// TIA Portal V19 export
VAR_GLOBAL   // PLC tag table "R3_IN"
   "ByteIN :0 R3" AT %IB154 : Byte;   // System Bits 1
   "ByteIN :1 R3" AT %IB155 : Byte;   // System Bits 2
   "ByteIN :2 R3" AT %IB156 : Byte;   // Signals
   "ByteIN :3 R3" AT %IB157 : Byte;   // Signals
   "ByteIN :4 R3" AT %IB158 : Byte;   // CMD
   "ByteIN :5 R3" AT %IB159 : Byte;
   "ByteIN :6 R3" AT %IB160 : Byte;
   "ByteIN :7 R3" AT %IB161 : Byte;
   "ByteIN :8 R3" AT %IB162 : Byte;
   "ByteIN :9 R3" AT %IB163 : Byte;
   "ByteIN :10 R3" AT %IB164 : Byte;
   "ByteIN :11 R3" AT %IB165 : Byte;
   "ByteIN :12 R3" AT %IB166 : Byte;
   "ByteIN :13 R3" AT %IB167 : Byte;
   "ByteIN :14 R3" AT %IB168 : Byte;
   "ByteIN :15 R3" AT %IB169 : Byte;
   "ByteIN :16 R3" AT %IB170 : Byte;
   "ByteIN :17 R3" AT %IB171 : Byte;
   "ByteIN :18 R3" AT %IB172 : Byte;
   "ByteIN :19 R3" AT %IB173 : Byte;
   "ByteIN :20 R3" AT %IB174 : Byte;
   "ByteIN :21 R3" AT %IB175 : Byte;
   "ByteIN :22 R3" AT %IB176 : Byte;
   "ByteIN :23 R3" AT %IB177 : Byte;
   "ByteIN :24 R3" AT %IB178 : Byte;
   "ByteIN :25 R3" AT %IB179 : Byte;
   "ByteIN :26 R3" AT %IB180 : Byte;
   "ByteIN :27 R3" AT %IB181 : Byte;
   "ByteIN :28 R3" AT %IB182 : Byte;
   "ByteIN :29 R3" AT %IB183 : Byte;
   "ByteIN :30 R3" AT %IB184 : Byte;
   "ByteIN :31 R3" AT %IB185 : Byte;
   "ByteIN :32 R3" AT %IB186 : Byte;
   "ByteIN :33 R3" AT %IB187 : Byte;
   "ByteIN :34 R3" AT %IB188 : Byte;
   "ByteIN :35 R3" AT %IB189 : Byte;
   "ByteIN :36 R3" AT %IB190 : Byte;
   "ByteIN :37 R3" AT %IB191 : Byte;
   "ByteIN :38 R3" AT %IB192 : Byte;
   "ByteIN :39 R3" AT %IB193 : Byte;
   "ByteIN :40 R3" AT %IB194 : Byte;
   "ByteIN :41 R3" AT %IB195 : Byte;
   "ByteIN :42 R3" AT %IB196 : Byte;
   "ByteIN :43 R3" AT %IB197 : Byte;
   "ByteIN :44 R3" AT %IB198 : Byte;
   "ByteIN :45 R3" AT %IB199 : Byte;
   "ByteIN :46 R3" AT %IB200 : Byte;
   "ByteIN :47 R3" AT %IB201 : Byte;
   "ByteIN :48 R3" AT %IB202 : Byte;
   "ByteIN :49 R3" AT %IB203 : Byte;
   "ByteIN :50 R3" AT %IB204 : Byte;
   "ByteIN :51 R3" AT %IB205 : Byte;
   "ByteIN :52 R3" AT %IB206 : Byte;
   "ByteIN :53 R3" AT %IB207 : Byte;
   "ByteIN :54 R3" AT %IB208 : Byte;
   "ByteIN :55 R3" AT %IB209 : Byte;
   "ByteIN :56 R3" AT %IB210 : Byte;
   "ByteIN :57 R3" AT %IB211 : Byte;
   "ByteIN :58 R3" AT %IB212 : Byte;
   "ByteIN :59 R3" AT %IB213 : Byte;
   "ByteIN :60 R3" AT %IB214 : Byte;
   "ByteIN :61 R3" AT %IB215 : Byte;
   "ByteIN :62 R3" AT %IB216 : Byte;
   "ByteIN :63 R3" AT %IB217 : Byte;
END_VAR
